(* IEC 61131-3 sources: plc-vscode/tests/st/all/trust-platform/examples/mitsubishi_gxworks3_v1/src, 2 files *)

(* ---- Main.st ---- *)
FUNCTION_BLOCK FB_EdgeBridge
VAR_INPUT
    Signal : BOOL;
END_VAR
VAR_OUTPUT
    Rising : BOOL;
    Falling : BOOL;
END_VAR
VAR
    UpEdge : DIFU;
    DownEdge : DIFD;
END_VAR

UpEdge(CLK := Signal, Q => Rising);
DownEdge(CLK := Signal, Q => Falling);
END_FUNCTION_BLOCK

PROGRAM Main
VAR
    Bridge : FB_EdgeBridge;
    Pulse : BOOL;
    RiseSeen : BOOL;
    FallSeen : BOOL;
END_VAR

Bridge(Signal := Pulse);
RiseSeen := Bridge.Rising;
FallSeen := Bridge.Falling;
END_PROGRAM

(* ---- Configuration.st ---- *)
CONFIGURATION MitsubishiDemo
RESOURCE MitsubishiRes ON PLC
TASK Cycle (INTERVAL := T#50ms, PRIORITY := 1);
PROGRAM P1 WITH Cycle : Main;
END_RESOURCE
VAR_CONFIG
    P1.Pulse AT %IX0.0 : BOOL;
    P1.RiseSeen AT %QX0.0 : BOOL;
    P1.FallSeen AT %QX0.1 : BOOL;
END_VAR
END_CONFIGURATION
